(* IEC 61131-3 sources: ZPLC/packages/zplc-ide/plant-scenes/height-sorting-chain, 2 files *)

(* ---- reference.st ---- *)
PROGRAM HeightSortChain
VAR_INPUT
    Start       AT %I0.0 : BOOL;
    Low         AT %I0.1 : BOOL;
    High        AT %I0.2 : BOOL;
    AtBlade     AT %I0.3 : BOOL;
    Raised      AT %I0.4 : BOOL;
    Lowered     AT %I0.5 : BOOL;
END_VAR
VAR_OUTPUT
    RunIn       AT %Q0.0 : BOOL;
    RunChain    AT %Q0.1 : BOOL;
    Lift        AT %Q0.2 : BOOL;
    MoveRight   AT %Q0.3 : BOOL;
    MoveLeft    AT %Q0.4 : BOOL;
    RunStraight AT %Q0.5 : BOOL;
    RunRight    AT %Q0.6 : BOOL;
    RunLeft     AT %Q0.7 : BOOL;
    Hold        AT %Q1.0 : BOOL;
    Busy        AT %Q1.1 : BOOL;
    Done        AT %Q1.2 : BOOL;
END_VAR
VAR
    Active   : BOOL;
    State    : INT;
    Dir      : INT;
    Handled  : INT;
    SawLow   : BOOL;
    SawHigh  : BOOL;
    Stand    : TON;
    Clear    : TON;
    Lifted   : TON;
    Slide    : TON;
END_VAR

IF Start THEN
    Active := TRUE;
END_IF;

(* the two beams sit across the infeed: 0.25 m (a 0.30 m or 0.40 m box breaks it) and 0.35 m (only
   a 0.40 m box breaks it). A 0.20 m box breaks neither. The latch keeps what the box showed. *)
IF Low THEN
    SawLow := TRUE;
END_IF;
IF High THEN
    SawHigh := TRUE;
END_IF;

(* the box must stand still against the blade before anything moves; the module needs a moment at the
   top before it slides a box (its surface stops first); the timers below are measured for 0.5 m/s *)
Stand(IN := AtBlade AND State = 1, PT := T#1000ms);
Clear(IN := State = 2, PT := T#2200ms);
Lifted(IN := State = 3 AND Raised, PT := T#300ms);
Slide(IN := State = 4, PT := T#1600ms);

(* 0 idle, 1 wait for a box at the blade, 2 straight on (short), 3 lift, 4 slide sideways, 5 lower.
   Dir: 0 short (straight), 1 medium (right), 2 tall (left) *)
CASE State OF
    0:
        IF Active THEN
            State := 1;
        END_IF;
    1:
        IF Stand.Q THEN
            IF SawHigh THEN
                Dir := 2;
            ELSIF SawLow THEN
                Dir := 1;
            ELSE
                Dir := 0;
            END_IF;
            (* the next box passes the beams before this one is done: clear the latch now *)
            SawLow := FALSE;
            SawHigh := FALSE;
            IF Dir = 0 THEN
                State := 2;
            ELSE
                State := 3;
            END_IF;
        END_IF;
    2:
        IF Clear.Q THEN
            Handled := Handled + 1;
            State := 1;
        END_IF;
    3:
        IF Lifted.Q THEN
            State := 4;
        END_IF;
    4:
        IF Slide.Q THEN
            State := 5;
        END_IF;
    5:
        IF Lowered THEN
            Handled := Handled + 1;
            State := 1;
        END_IF;
END_CASE;

RunIn       := Active;
RunStraight := Active;
RunRight    := Active;
RunLeft     := Active;
(* the module carries a box straight on while it is down; with lift it must not run (a conflict) *)
RunChain    := Active AND (State = 1 OR State = 2);
Hold        := Active AND State <> 2;
Lift        := State = 3 OR State = 4;
MoveRight   := State = 4 AND Dir = 1;
MoveLeft    := State = 4 AND Dir = 2;
Busy        := Active AND Handled < 9;
Done        := Handled >= 9;

END_PROGRAM

(* ---- starter.st ---- *)
PROGRAM HeightSortChain
VAR_INPUT
    Start       AT %I0.0 : BOOL;  (* StartButton.pressed: start the line *)
    Low         AT %I0.1 : BOOL;  (* BeamLow.detect: a box 0.30 m or 0.40 m high breaks the lower beam *)
    High        AT %I0.2 : BOOL;  (* BeamHigh.detect: a box 0.40 m high breaks the upper beam *)
    AtBlade     AT %I0.3 : BOOL;  (* EyeChain.detect: a box stands against the blade on the transfer *)
    Raised      AT %I0.4 : BOOL;  (* Chain1.raised: the chain module is up *)
    Lowered     AT %I0.5 : BOOL;  (* Chain1.lowered: the chain module is down *)
END_VAR
VAR_OUTPUT
    RunIn       AT %Q0.0 : BOOL;  (* Infeed.run: run the infeed belt *)
    RunChain    AT %Q0.1 : BOOL;  (* Chain1.run: run the module straight on while it is down *)
    Lift        AT %Q0.2 : BOOL;  (* Chain1.lift: raise the module while true *)
    MoveRight   AT %Q0.3 : BOOL;  (* Chain1.moveRight: move a box to the right belt (module up) *)
    MoveLeft    AT %Q0.4 : BOOL;  (* Chain1.moveLeft: move a box to the left belt (module up) *)
    RunStraight AT %Q0.5 : BOOL;  (* Straight.run: run the belt beyond the transfer *)
    RunRight    AT %Q0.6 : BOOL;  (* SideRight.run: run the right belt *)
    RunLeft     AT %Q0.7 : BOOL;  (* SideLeft.run: run the left belt *)
    Hold        AT %Q1.0 : BOOL;  (* Stop1.extend: the blade holds a box on the module while true *)
    Busy        AT %Q1.1 : BOOL;  (* Beacon.amber: the line is running *)
    Done        AT %Q1.2 : BOOL;  (* Beacon.green: lit when nine boxes have been sorted *)
END_VAR

(* Goal: a press of the start button runs every belt. Boxes of three heights (0.20, 0.30 and
   0.40 m) arrive on the infeed, one every five seconds, nine in all. Tell the height from the
   two beams while the box passes them: 0.20 m breaks neither, 0.30 m only the lower, 0.40 m both.
   Remember the answer, because the box reaches the transfer later and the next box may pass the
   beams before this one is done.
   A box stops against the blade on the chain module (hold the blade, and run the module so that
   the box is pushed against it). Once it has stood still for a second:
     - 0.20 m: release the blade and run the module; the box goes straight on to the short bin;
     - 0.30 m: stop the module, lift it, wait until it is up and has rested a moment, then move
       right until the box is on the right belt, and lower the module (medium bin);
     - 0.40 m: the same, to the left (tall bin).
   Never run the module and lift it at the same time. Light Busy while the line runs and Done when
   nine boxes have been sorted. *)

END_PROGRAM
